// TIA Portal V21 export
VAR_GLOBAL   // PLC tag table "StateConstant"
END_VAR
VAR_GLOBAL CONSTANT   // user constants
   ST3_AUTOMATIC_INIT : Int := 3;
   ST999_FAULT : Int := 999;
   ST1_READY : Int := 1;
   ST2_STARTING : Int := 2;
   ST4_AUTOMATIC_PAUSE : Int := 4;
   ST5_SHUTDOWN : Int := 5;
   ST900_QUICKSTOP : Int := 900;
   ST0_STOPPED : Int := 0;
END_VAR
